// TIA Portal project "TIA_KONE_MOHAMED_EXERCICE1" (V16)

(* hardware
DEVICE "Station S7300/ET200M_1"  S7-300 station
   slot 0: "Châssis_0"  Rail  6ES7 390-1***0-0AA0
   slot 2: "PLC_1"  CPU 313C  6ES7 313-5BG04-0AB0  V3.3
      slot 0: "Interface MPI_1"  MPI
      slot 2: "DI 24/DO 16_1"  DI24/DO16
      slot 3: "AI 5/AO 2_1"  AI5/AO2
      slot 4: "Comptage_1"  Counter
*)

// ===== PLC "PLC_1"  CPU 313C =====

VAR_GLOBAL   // PLC tag table "Table de variables standard"
   "X31" AT %Q1.4 : Bool;
   "a0" AT %I0.1 : Bool;
   "b1" AT %I0.4 : Bool;
   "X41" AT %Q1.5 : Bool;
   "X1" AT %Q1.0 : Bool;
   "X2" AT %Q1.1 : Bool;
   "X30" AT %Q1.2 : Bool;
   "X40" AT %Q1.3 : Bool;
   "DCY" AT %I0.0 : Bool;
   "tr" AT %I0.6 : Bool;
   "Pr" AT %I0.7 : Bool;
   "a1" AT %I0.2 : Bool;
   "b0" AT %I0.3 : Bool;
   "KM1" AT %Q0.0 : Bool;
   "A+" AT %Q0.1 : Bool;
   "A-" AT %Q0.2 : Bool;
   "B-" AT %Q0.4 : Bool;
   "B+" AT %Q0.3 : Bool;
   "MARCHE" AT %I2.1 : Bool;
   "M" AT %M2.2 : Bool;
END_VAR

ORGANIZATION_BLOCK "Main"   // OB1, LAD
TITLE = "Main Program Sweep (Cycle)"
{ S7_Optimized_Access := 'FALSE' }
VERSION : 0.1
   VAR_TEMP
      OB1_EV_CLASS : Byte;   // Bits 0-3 = 1 (Coming event), Bits 4-7 = 1 (Event class 1)
      OB1_SCAN_1 : Byte;   // 1 (Cold restart scan 1 of OB 1), 3 (Scan 2-n of OB 1)
      OB1_PRIORITY : Byte;   // Priority of OB Execution
      OB1_OB_NUMBR : Byte;   // 1 (Organization block 1, OB1)
      OB1_RESERVED_1 : Byte;   // Reserved for system
      OB1_RESERVED_2 : Byte;   // Reserved for system
      OB1_PREV_CYCLE : Int;   // Cycle time of previous OB1 scan (milliseconds)
      OB1_MIN_CYCLE : Int;   // Minimum cycle time of OB1 (milliseconds)
      OB1_MAX_CYCLE : Int;   // Maximum cycle time of OB1 (milliseconds)
      OB1_DATE_TIME : Date_And_Time;   // Date and time OB1 started
   END_VAR
   VAR_TEMP   // added for the SCL form of the ladder/FBD networks
      _w1 : Bool;
   END_VAR
BEGIN

REGION Network 1
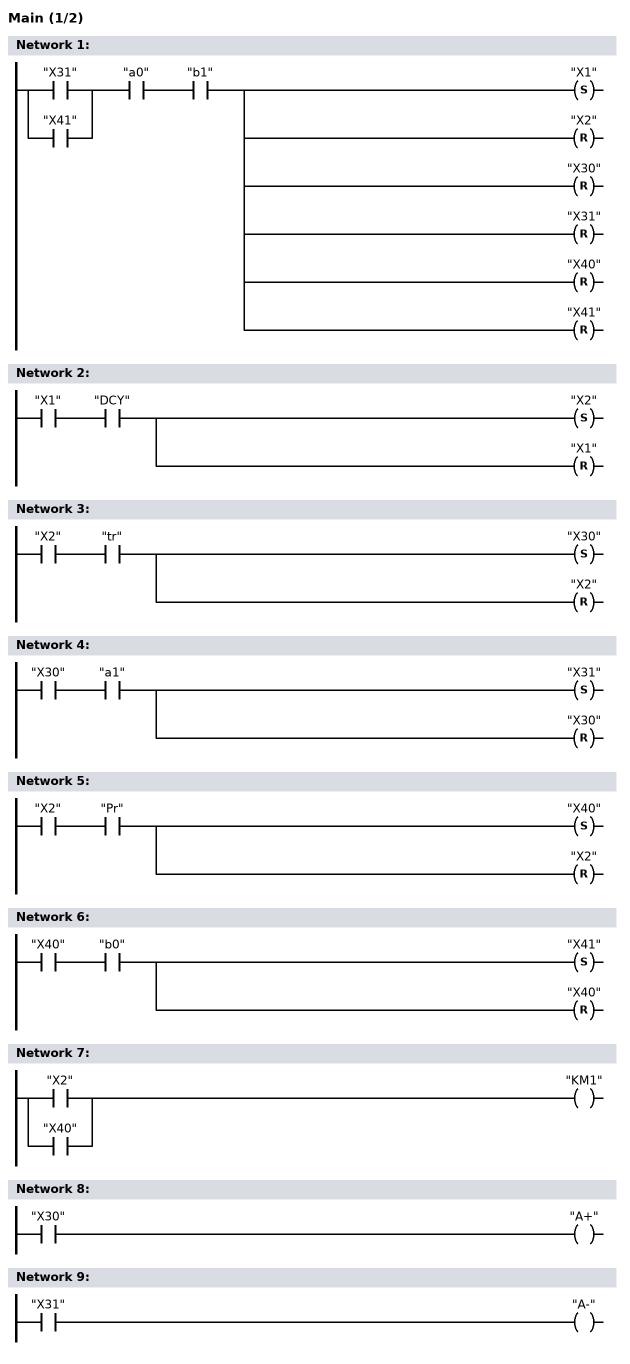
   RUNG wire#powerrail
      Contact( "X31" )
      wire#w1
      Contact( "a0" )
      Contact( "b1" )
      wire#w2
      S_Coil( "X1" )
   END_RUNG
   RUNG wire#powerrail
      Contact( "X41" )
   END_RUNG wire#w1
   RUNG wire#w2
      R_Coil( "X2" )
   END_RUNG
   RUNG wire#w2
      R_Coil( "X30" )
   END_RUNG
   RUNG wire#w2
      R_Coil( "X31" )
   END_RUNG
   RUNG wire#w2
      R_Coil( "X40" )
   END_RUNG
   RUNG wire#w2
      R_Coil( "X41" )
   END_RUNG
   // the same network as SCL:
   IF ("X31" OR "X41") AND "a0" AND "b1" THEN
       "X1" := TRUE;
       "X2" := FALSE;
       "X30" := FALSE;
   END_IF;
   #_w1 := ("X31" OR "X41") AND "a0" AND "b1";
   IF #_w1 THEN
       "X31" := FALSE;
       "X40" := FALSE;
       "X41" := FALSE;
   END_IF;
END_REGION

REGION Network 2
   RUNG wire#powerrail
      Contact( "X1" )
      Contact( "DCY" )
      wire#w1
      S_Coil( "X2" )
   END_RUNG
   RUNG wire#w1
      R_Coil( "X1" )
   END_RUNG
   // the same network as SCL:
   IF "X1" AND "DCY" THEN
       "X2" := TRUE;
       "X1" := FALSE;
   END_IF;
END_REGION

REGION Network 3
   RUNG wire#powerrail
      Contact( "X2" )
      Contact( "tr" )
      wire#w1
      S_Coil( "X30" )
   END_RUNG
   RUNG wire#w1
      R_Coil( "X2" )
   END_RUNG
   // the same network as SCL:
   IF "X2" AND "tr" THEN
       "X30" := TRUE;
       "X2" := FALSE;
   END_IF;
END_REGION

REGION Network 4
   RUNG wire#powerrail
      Contact( "X30" )
      Contact( "a1" )
      wire#w1
      S_Coil( "X31" )
   END_RUNG
   RUNG wire#w1
      R_Coil( "X30" )
   END_RUNG
   // the same network as SCL:
   IF "X30" AND "a1" THEN
       "X31" := TRUE;
       "X30" := FALSE;
   END_IF;
END_REGION

REGION Network 5
   RUNG wire#powerrail
      Contact( "X2" )
      Contact( "Pr" )
      wire#w1
      S_Coil( "X40" )
   END_RUNG
   RUNG wire#w1
      R_Coil( "X2" )
   END_RUNG
   // the same network as SCL:
   IF "X2" AND "Pr" THEN
       "X40" := TRUE;
       "X2" := FALSE;
   END_IF;
END_REGION

REGION Network 6
   RUNG wire#powerrail
      Contact( "X40" )
      Contact( "b0" )
      wire#w1
      S_Coil( "X41" )
   END_RUNG
   RUNG wire#w1
      R_Coil( "X40" )
   END_RUNG
   // the same network as SCL:
   IF "X40" AND "b0" THEN
       "X41" := TRUE;
       "X40" := FALSE;
   END_IF;
END_REGION

REGION Network 7
   RUNG wire#powerrail
      Contact( "X2" )
      wire#w1
      Coil( "KM1" )
   END_RUNG
   RUNG wire#powerrail
      Contact( "X40" )
   END_RUNG wire#w1
   // the same network as SCL:
   "KM1" := "X2" OR "X40";
END_REGION

REGION Network 8
   RUNG wire#powerrail
      Contact( "X30" )
      Coil( "A+" )
   END_RUNG
   // the same network as SCL:
   "A+" := "X30";
END_REGION

REGION Network 9
   RUNG wire#powerrail
      Contact( "X31" )
      Coil( "A-" )
   END_RUNG
   // the same network as SCL:
   "A-" := "X31";
END_REGION

REGION Network 10
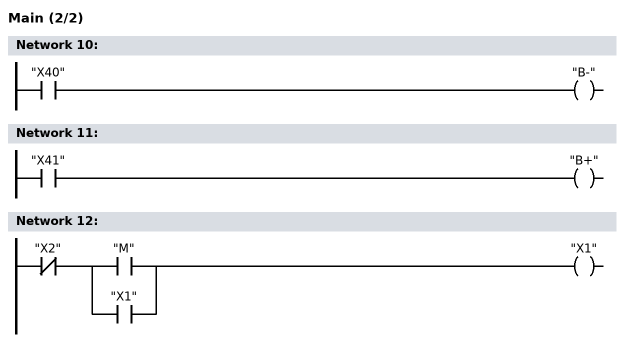
   RUNG wire#powerrail
      Contact( "X40" )
      Coil( "B-" )
   END_RUNG
   // the same network as SCL:
   "B-" := "X40";
END_REGION

REGION Network 11
   RUNG wire#powerrail
      Contact( "X41" )
      Coil( "B+" )
   END_RUNG
   // the same network as SCL:
   "B+" := "X41";
END_REGION

REGION Network 12
   RUNG wire#powerrail
      I_Contact( "X2" )
      wire#w1
      Contact( "M" )
      wire#w2
      Coil( "X1" )
   END_RUNG
   RUNG wire#w1
      Contact( "X1" )
   END_RUNG wire#w2
   // the same network as SCL:
   "X1" := NOT "X2" AND ("M" OR "X1");
END_REGION
END_ORGANIZATION_BLOCK